//---------------------------------------------------------------------------------------------------------------
//
//  HAUD 2026.10.25
//
//  - ExternControl
//
//    - this is the main switchboard
//
//    - Transport abstractions are called here:
//    --------------------------------------------
//    - top level transport abstractions
//      - Instances contain the required transport logic
//      - Instances control their assigned ProcessCollector
//      - Instances are controlled in timer based application
//
//    - mid level transport abstractions
//      - StationCollectors and by extension ProcessCollectors
//      - Collectors are for gathering states and routing commands to ST_STATION_CTRL/STATE
//      - Collectors are configured during startup
//
//---------------------------------------------------------------------------------------------------------------
PROGRAM MAIN_APP
VAR
  eInitXtsTransport   AT %I*    : E_PROGRESS;   // initialization from XtsTransport PLC
  eInit               AT %Q*    : E_PROGRESS;   // local startup transmitted to TowerControl

  idx                           : UINT;
  nProcess                      : E_INSTANCE;

  // message pipeline(s) handling
  eMtrState,
  eMsgState                     : E_MESSAGE_STATE;
  eMtrProgress,
  eMsgProgress                  : E_PROGRESS;
  stMsg                         : ST_Message;
  //-------------------------------------------------------------------------------------------------------------
  tIdleWriteMotion              : TIME := T#5S;
  tIdleWriteApplication         : TIME := T#5S;
  tIdleWriteMetric              : TIME := T#5S;
  tonIdleWriteMotion            : Tc2_Standard.TON;
  tonIdleWriteApplication       : Tc2_Standard.TON;
  tonIdleWriteMetric            : Tc2_Standard.TON;
  //-------------------------------------------------------------------------------------------------------------
END_VAR

//#################################################################################################################
// Local time; used for timestamps
//#################################################################################################################
GVL_MSG_XTS.fbLocalTime();
GVL_MSG_XTS.sLocalTime                                            := GVL_MSG_XTS.fbLocalTime.LocalTimeString;
GVL_MSG_XTS.dtLocalTime                                           := GVL_MSG_XTS.fbLocalTime.LocalTime;
//-----------------------------------------------------------------------------------------------------------------
//-----------------------------------------------------------------------------------------------------------------
// check for Initialisation from XtsTransport first
//  - wait for XtsTransport to be fully started up
//-----------------------------------------------------------------------------------------------------------------
IF NOT (eInitXtsTransport = E_PROGRESS.PROGRESS_DONE) THEN eInit  := E_PROGRESS.PROGRESS_INVALID; RETURN; END_IF
//-----------------------------------------------------------------------------------------------------------------
//-----------------------------------------------------------------------------------------------------------------
// initialization for:
//  - configuring processes
//  - starting up of processes
//  - cross checking with the rest of your application
//-----------------------------------------------------------------------------------------------------------------
CASE eInit
OF
  E_PROGRESS.PROGRESS_INVALID:
    GVL_MSG_XTS.MetricsMessageCtrl.Cmd            := E_MESSAGE_CTRL.MSG_CTRL_INIT;
    eInit                                         := E_PROGRESS.PROGRESS_INIT;

  E_PROGRESS.PROGRESS_INIT:
    // init processes
    eInit                                         := E_PROGRESS.PROGRESS_BUSY;
    //-----------------------------------------------------------------------------
    //#############################################################################
    //-----------------------------------------------------------------------------
    GVL_APPLICATION.ProcessCollector[DISTRIBUTOR_INFEED].ProcessId            := DISTRIBUTOR_INFEED;
    GVL_APPLICATION.ProcessCollector[DISTRIBUTOR_INFEED].StationFirst         :=   142;
    GVL_APPLICATION.ProcessCollector[DISTRIBUTOR_INFEED].StationLast          :=   142;
    //-----------------------------------------------------------------------------
    GVL_APPLICATION.InstanceDistributorInfeed.ProcessId                       := DISTRIBUTOR_INFEED;
    GVL_APPLICATION.InstanceDistributorInfeed.ProcessTarget                   := PROCESS_INFEED;
    GVL_APPLICATION.InstanceDistributorInfeed.CheckPositionStart              :=  4500.0;
    GVL_APPLICATION.InstanceDistributorInfeed.CheckPositionEnd                :=  5600.0;
    //-----------------------------------------------------------------------------
    GVL_APPLICATION.InstanceDistributorInfeed.CollectorInterface              :=   GVL_APPLICATION.ItfProcessCollector;
    GVL_APPLICATION.InstanceDistributorInfeed.ProcessLinkedLists              :=   GVL_APPLICATION.ItfProcessList;
    GVL_APPLICATION.InstanceDistributorInfeed.InstanceCtrl                    REF= GVL_APPLICATION.InstanceCtrl;
    GVL_APPLICATION.InstanceDistributorInfeed.InstanceState                   REF= GVL_APPLICATION.InstanceState;
    GVL_APPLICATION.InstanceDistributorInfeed.MessageLevel                    :=   E_MessageType.eMessageError;

    //-----------------------------------------------------------------------------
    //#############################################################################
    //-----------------------------------------------------------------------------
    GVL_APPLICATION.ProcessCollector[PROCESS_INFEED].ProcessId                := PROCESS_INFEED;
    GVL_APPLICATION.ProcessCollector[PROCESS_INFEED].StationFirst             :=    20;
    GVL_APPLICATION.ProcessCollector[PROCESS_INFEED].StationLast              :=    35;
    //-----------------------------------------------------------------------------
    GVL_APPLICATION.InstanceInfeed.ProcessId                                  := PROCESS_INFEED;
    GVL_APPLICATION.InstanceInfeed.ProcessTarget                              := CONTINUOUS_CLEAN;
    GVL_APPLICATION.InstanceInfeed.CheckPositionStart                         :=  9750.0;
    GVL_APPLICATION.InstanceInfeed.CheckPositionEnd                           := 12100.0;
    //-----------------------------------------------------------------------------
    GVL_APPLICATION.InstanceInfeed.CollectorInterface                         :=   GVL_APPLICATION.ItfProcessCollector;
    GVL_APPLICATION.InstanceInfeed.ProcessLinkedLists                         :=   GVL_APPLICATION.ItfProcessList;
    GVL_APPLICATION.InstanceInfeed.InstanceCtrl                               REF= GVL_APPLICATION.InstanceCtrl;
    GVL_APPLICATION.InstanceInfeed.InstanceState                              REF= GVL_APPLICATION.InstanceState;
    GVL_APPLICATION.InstanceInfeed.MessageLevel                               :=   E_MessageType.eMessageError;

    //-----------------------------------------------------------------------------
    //#############################################################################
    //-----------------------------------------------------------------------------
    GVL_APPLICATION.ProcessCollector[CONTINUOUS_CLEAN].ProcessId              := CONTINUOUS_CLEAN;
    GVL_APPLICATION.ProcessCollector[CONTINUOUS_CLEAN].StationFirst           :=    37;
    GVL_APPLICATION.ProcessCollector[CONTINUOUS_CLEAN].StationLast            :=    37;
    //-----------------------------------------------------------------------------
    GVL_APPLICATION.InstanceCleaner.ProcessId                                 := CONTINUOUS_CLEAN;
    GVL_APPLICATION.InstanceCleaner.ProcessTarget                             := CONTINUOUS_SCAN;
    GVL_APPLICATION.InstanceCleaner.CheckPositionStart                        := 12850.0;
    GVL_APPLICATION.InstanceCleaner.CheckPositionEnd                          := 13000.0;
    //-----------------------------------------------------------------------------
    GVL_APPLICATION.InstanceCleaner.CollectorInterface                        :=   GVL_APPLICATION.ItfProcessCollector;
    GVL_APPLICATION.InstanceCleaner.ProcessLinkedLists                        :=   GVL_APPLICATION.ItfProcessList;
    GVL_APPLICATION.InstanceCleaner.InstanceCtrl                              REF= GVL_APPLICATION.InstanceCtrl;
    GVL_APPLICATION.InstanceCleaner.InstanceState                             REF= GVL_APPLICATION.InstanceState;

    //-----------------------------------------------------------------------------
    //#############################################################################
    //-----------------------------------------------------------------------------
    GVL_APPLICATION.ProcessCollector[CONTINUOUS_SCAN].ProcessId               := CONTINUOUS_SCAN;
    GVL_APPLICATION.ProcessCollector[CONTINUOUS_SCAN].StationFirst            :=    38;
    GVL_APPLICATION.ProcessCollector[CONTINUOUS_SCAN].StationLast             :=    38;
    //-----------------------------------------------------------------------------
    GVL_APPLICATION.InstanceScanner.ProcessId                                 := CONTINUOUS_SCAN;
    GVL_APPLICATION.InstanceScanner.ProcessTarget                             := CONTINUOUS_CAMERA;
    GVL_APPLICATION.InstanceScanner.CheckPositionStart                        := 13900.0;
    GVL_APPLICATION.InstanceScanner.CheckPositionEnd                          := 14100.0;
    //-----------------------------------------------------------------------------
    GVL_APPLICATION.InstanceScanner.CollectorInterface                        :=   GVL_APPLICATION.ItfProcessCollector;
    GVL_APPLICATION.InstanceScanner.ProcessLinkedLists                        :=   GVL_APPLICATION.ItfProcessList;
    GVL_APPLICATION.InstanceScanner.InstanceCtrl                              REF= GVL_APPLICATION.InstanceCtrl;
    GVL_APPLICATION.InstanceScanner.InstanceState                             REF= GVL_APPLICATION.InstanceState;

    //-----------------------------------------------------------------------------
    //#############################################################################
    //-----------------------------------------------------------------------------
    GVL_APPLICATION.ProcessCollector[CONTINUOUS_CAMERA].ProcessId             := CONTINUOUS_CAMERA;
    GVL_APPLICATION.ProcessCollector[CONTINUOUS_CAMERA].StationFirst          :=    39;
    GVL_APPLICATION.ProcessCollector[CONTINUOUS_CAMERA].StationLast           :=    39;
    //-----------------------------------------------------------------------------
    GVL_APPLICATION.InstanceCamera.ProcessId                                  := CONTINUOUS_CAMERA;
    GVL_APPLICATION.InstanceCamera.ProcessTarget                              := DISTRIBUTOR_ASSEMBLY_01;
    GVL_APPLICATION.InstanceCamera.CheckPositionStart                         := 14200.0;
    GVL_APPLICATION.InstanceCamera.CheckPositionEnd                           := 14400.0;
    //-----------------------------------------------------------------------------
    GVL_APPLICATION.InstanceCamera.CollectorInterface                         :=   GVL_APPLICATION.ItfProcessCollector;
    GVL_APPLICATION.InstanceCamera.ProcessLinkedLists                         :=   GVL_APPLICATION.ItfProcessList;
    GVL_APPLICATION.InstanceCamera.InstanceCtrl                               REF= GVL_APPLICATION.InstanceCtrl;
    GVL_APPLICATION.InstanceCamera.InstanceState                              REF= GVL_APPLICATION.InstanceState;

    //-----------------------------------------------------------------------------
    //#############################################################################
    //-----------------------------------------------------------------------------
    GVL_APPLICATION.ProcessCollector[DISTRIBUTOR_ASSEMBLY_01].ProcessId       := DISTRIBUTOR_ASSEMBLY_01;
    GVL_APPLICATION.ProcessCollector[DISTRIBUTOR_ASSEMBLY_01].StationFirst    :=    40;
    GVL_APPLICATION.ProcessCollector[DISTRIBUTOR_ASSEMBLY_01].StationLast     :=    40;
    //-----------------------------------------------------------------------------
    GVL_APPLICATION.InstanceDistributorAssembly_01.ProcessId                  := DISTRIBUTOR_ASSEMBLY_01;
    GVL_APPLICATION.InstanceDistributorAssembly_01.ProcessTarget              := PROCESS_ASSEMBLY_01;
    GVL_APPLICATION.InstanceDistributorAssembly_01.CheckPositionStart         := 14400.0;
    GVL_APPLICATION.InstanceDistributorAssembly_01.CheckPositionEnd           := 17500.0;
    //-----------------------------------------------------------------------------
    GVL_APPLICATION.InstanceDistributorAssembly_01.CollectorInterface         :=   GVL_APPLICATION.ItfProcessCollector;
    GVL_APPLICATION.InstanceDistributorAssembly_01.ProcessLinkedLists         :=   GVL_APPLICATION.ItfProcessList;
    GVL_APPLICATION.InstanceDistributorAssembly_01.InstanceCtrl               REF= GVL_APPLICATION.InstanceCtrl;
    GVL_APPLICATION.InstanceDistributorAssembly_01.InstanceState              REF= GVL_APPLICATION.InstanceState;

    //-----------------------------------------------------------------------------
    //#############################################################################
    //-----------------------------------------------------------------------------
    GVL_APPLICATION.ProcessCollector[PROCESS_ASSEMBLY_01].ProcessId           := PROCESS_ASSEMBLY_01;
    GVL_APPLICATION.ProcessCollector[PROCESS_ASSEMBLY_01].StationFirst        :=    41;
    GVL_APPLICATION.ProcessCollector[PROCESS_ASSEMBLY_01].StationLast         :=    56;
    //-----------------------------------------------------------------------------
    GVL_APPLICATION.InstanceAssembly_01.ProcessId                             := PROCESS_ASSEMBLY_01;
    GVL_APPLICATION.InstanceAssembly_01.ProcessTarget                         := DISTRIBUTOR_ASSEMBLY_02;
    GVL_APPLICATION.InstanceAssembly_01.CheckPositionStart                    := 14400.0;
    GVL_APPLICATION.InstanceAssembly_01.CheckPositionEnd                      := 17500.0;
    //-----------------------------------------------------------------------------
    GVL_APPLICATION.InstanceAssembly_01.CollectorInterface                    :=   GVL_APPLICATION.ItfProcessCollector;
    GVL_APPLICATION.InstanceAssembly_01.ProcessLinkedLists                    :=   GVL_APPLICATION.ItfProcessList;
    GVL_APPLICATION.InstanceAssembly_01.InstanceCtrl                          REF= GVL_APPLICATION.InstanceCtrl;
    GVL_APPLICATION.InstanceAssembly_01.InstanceState                         REF= GVL_APPLICATION.InstanceState;

    //-----------------------------------------------------------------------------
    //#############################################################################
    //-----------------------------------------------------------------------------
    GVL_APPLICATION.ProcessCollector[DISTRIBUTOR_ASSEMBLY_02].ProcessId       := DISTRIBUTOR_ASSEMBLY_02;
    GVL_APPLICATION.ProcessCollector[DISTRIBUTOR_ASSEMBLY_02].StationFirst    :=    57;
    GVL_APPLICATION.ProcessCollector[DISTRIBUTOR_ASSEMBLY_02].StationLast     :=    57;
    //-----------------------------------------------------------------------------
    GVL_APPLICATION.InstanceDistributorAssembly_02.ProcessId                  := DISTRIBUTOR_ASSEMBLY_02;
    GVL_APPLICATION.InstanceDistributorAssembly_02.ProcessTarget              := PROCESS_ASSEMBLY_02;
    GVL_APPLICATION.InstanceDistributorAssembly_02.CheckPositionStart         := 17500.0;
    GVL_APPLICATION.InstanceDistributorAssembly_02.CheckPositionEnd           := 18100.0;
    //-----------------------------------------------------------------------------
    GVL_APPLICATION.InstanceDistributorAssembly_02.CollectorInterface         :=   GVL_APPLICATION.ItfProcessCollector;
    GVL_APPLICATION.InstanceDistributorAssembly_02.ProcessLinkedLists         :=   GVL_APPLICATION.ItfProcessList;
    GVL_APPLICATION.InstanceDistributorAssembly_02.InstanceCtrl               REF= GVL_APPLICATION.InstanceCtrl;
    GVL_APPLICATION.InstanceDistributorAssembly_02.InstanceState              REF= GVL_APPLICATION.InstanceState;

    //-----------------------------------------------------------------------------
    //#############################################################################
    //-----------------------------------------------------------------------------
    GVL_APPLICATION.ProcessCollector[PROCESS_ASSEMBLY_02].ProcessId           := PROCESS_ASSEMBLY_02;
    GVL_APPLICATION.ProcessCollector[PROCESS_ASSEMBLY_02].StationFirst        :=    58;
    GVL_APPLICATION.ProcessCollector[PROCESS_ASSEMBLY_02].StationLast         :=    67;
    //-----------------------------------------------------------------------------
    GVL_APPLICATION.InstanceAssembly_02.ProcessId                             := PROCESS_ASSEMBLY_02;
    GVL_APPLICATION.InstanceAssembly_02.ProcessTarget                         := DISTRIBUTOR_ASSEMBLY_TEST;
    GVL_APPLICATION.InstanceAssembly_02.CheckPositionStart                    := 19400.0;
    GVL_APPLICATION.InstanceAssembly_02.CheckPositionEnd                      := 20750.0;
    //-----------------------------------------------------------------------------
    GVL_APPLICATION.InstanceAssembly_02.CollectorInterface                    :=   GVL_APPLICATION.ItfProcessCollector;
    GVL_APPLICATION.InstanceAssembly_02.ProcessLinkedLists                    :=   GVL_APPLICATION.ItfProcessList;
    GVL_APPLICATION.InstanceAssembly_02.InstanceCtrl                          REF= GVL_APPLICATION.InstanceCtrl;
    GVL_APPLICATION.InstanceAssembly_02.InstanceState                         REF= GVL_APPLICATION.InstanceState;

    //-----------------------------------------------------------------------------
    //#############################################################################
    //-----------------------------------------------------------------------------
    GVL_APPLICATION.ProcessCollector[DISTRIBUTOR_ASSEMBLY_TEST].ProcessId     := DISTRIBUTOR_ASSEMBLY_TEST;
    GVL_APPLICATION.ProcessCollector[DISTRIBUTOR_ASSEMBLY_TEST].StationFirst  :=    70;
    GVL_APPLICATION.ProcessCollector[DISTRIBUTOR_ASSEMBLY_TEST].StationLast   :=    70;
    //-----------------------------------------------------------------------------
    GVL_APPLICATION.InstanceDistributorAssemblyTest.ProcessId                 := DISTRIBUTOR_ASSEMBLY_TEST;
    GVL_APPLICATION.InstanceDistributorAssemblyTest.ProcessTarget             := PROCESS_ASSEMBLY_TEST;
    GVL_APPLICATION.InstanceDistributorAssemblyTest.CheckPositionStart        := 20600.0;
    GVL_APPLICATION.InstanceDistributorAssemblyTest.CheckPositionEnd          := 21400.0;
    //-----------------------------------------------------------------------------
    GVL_APPLICATION.InstanceDistributorAssemblyTest.CollectorInterface        :=   GVL_APPLICATION.ItfProcessCollector;
    GVL_APPLICATION.InstanceDistributorAssemblyTest.ProcessLinkedLists        :=   GVL_APPLICATION.ItfProcessList;
    GVL_APPLICATION.InstanceDistributorAssemblyTest.InstanceCtrl              REF= GVL_APPLICATION.InstanceCtrl;
    GVL_APPLICATION.InstanceDistributorAssemblyTest.InstanceState             REF= GVL_APPLICATION.InstanceState;

    //-----------------------------------------------------------------------------
    //#############################################################################
    //-----------------------------------------------------------------------------
    GVL_APPLICATION.ProcessCollector[PROCESS_ASSEMBLY_TEST].ProcessId         := PROCESS_ASSEMBLY_TEST;
    GVL_APPLICATION.ProcessCollector[PROCESS_ASSEMBLY_TEST].StationFirst      :=    71;
    GVL_APPLICATION.ProcessCollector[PROCESS_ASSEMBLY_TEST].StationLast       :=    86;
    //-----------------------------------------------------------------------------
    GVL_APPLICATION.InstanceAssemblyTest.ProcessId                            := PROCESS_ASSEMBLY_TEST;
    GVL_APPLICATION.InstanceAssemblyTest.ProcessTarget                        := DISTRIBUTOR_CAMERA;
    GVL_APPLICATION.InstanceAssemblyTest.CheckPositionStart                   := 21400.0;
    GVL_APPLICATION.InstanceAssemblyTest.CheckPositionEnd                     := 23000.0;
    //-----------------------------------------------------------------------------
    GVL_APPLICATION.InstanceAssemblyTest.CollectorInterface                   :=   GVL_APPLICATION.ItfProcessCollector;
    GVL_APPLICATION.InstanceAssemblyTest.ProcessLinkedLists                   :=   GVL_APPLICATION.ItfProcessList;
    GVL_APPLICATION.InstanceAssemblyTest.InstanceCtrl                         REF= GVL_APPLICATION.InstanceCtrl;
    GVL_APPLICATION.InstanceAssemblyTest.InstanceState                        REF= GVL_APPLICATION.InstanceState;

    //-----------------------------------------------------------------------------
    //#############################################################################
    //-----------------------------------------------------------------------------
    GVL_APPLICATION.ProcessCollector[DISTRIBUTOR_CAMERA].ProcessId            := DISTRIBUTOR_CAMERA;
    GVL_APPLICATION.ProcessCollector[DISTRIBUTOR_CAMERA].StationFirst         :=    91;
    GVL_APPLICATION.ProcessCollector[DISTRIBUTOR_CAMERA].StationLast          :=    91;
    //-----------------------------------------------------------------------------
    GVL_APPLICATION.InstanceAssemblyCameraInfeed.ProcessId                    := DISTRIBUTOR_CAMERA;
    GVL_APPLICATION.InstanceAssemblyCameraInfeed.ProcessTarget                := CONTINUOUS_ASSEMBLY_CAMERA;
    GVL_APPLICATION.InstanceAssemblyCameraInfeed.CheckPositionStart           := 22800.0;
    GVL_APPLICATION.InstanceAssemblyCameraInfeed.CheckPositionEnd             := 23500.0;
    //-----------------------------------------------------------------------------
    GVL_APPLICATION.InstanceAssemblyCameraInfeed.CollectorInterface           :=   GVL_APPLICATION.ItfProcessCollector;
    GVL_APPLICATION.InstanceAssemblyCameraInfeed.ProcessLinkedLists           :=   GVL_APPLICATION.ItfProcessList;
    GVL_APPLICATION.InstanceAssemblyCameraInfeed.InstanceCtrl                 REF= GVL_APPLICATION.InstanceCtrl;
    GVL_APPLICATION.InstanceAssemblyCameraInfeed.InstanceState                REF= GVL_APPLICATION.InstanceState;

    //-----------------------------------------------------------------------------
    //#############################################################################
    //-----------------------------------------------------------------------------
    GVL_APPLICATION.ProcessCollector[CONTINUOUS_ASSEMBLY_CAMERA].ProcessId    := CONTINUOUS_ASSEMBLY_CAMERA;
    GVL_APPLICATION.ProcessCollector[CONTINUOUS_ASSEMBLY_CAMERA].StationFirst :=    95;
    GVL_APPLICATION.ProcessCollector[CONTINUOUS_ASSEMBLY_CAMERA].StationLast  :=    95;
    //-----------------------------------------------------------------------------
    GVL_APPLICATION.InstanceAssemblyCameraOutfeed.ProcessId                   := CONTINUOUS_ASSEMBLY_CAMERA;
    GVL_APPLICATION.InstanceAssemblyCameraOutfeed.ProcessTarget               := DISTRIBUTOR_OUTFEED;
    GVL_APPLICATION.InstanceAssemblyCameraOutfeed.CheckPositionStart          := 24000.0;
    GVL_APPLICATION.InstanceAssemblyCameraOutfeed.CheckPositionEnd            := 24100.0;
    //-----------------------------------------------------------------------------
    GVL_APPLICATION.InstanceAssemblyCameraOutfeed.CollectorInterface          :=   GVL_APPLICATION.ItfProcessCollector;
    GVL_APPLICATION.InstanceAssemblyCameraOutfeed.ProcessLinkedLists          :=   GVL_APPLICATION.ItfProcessList;
    GVL_APPLICATION.InstanceAssemblyCameraOutfeed.InstanceCtrl                REF= GVL_APPLICATION.InstanceCtrl;
    GVL_APPLICATION.InstanceAssemblyCameraOutfeed.InstanceState               REF= GVL_APPLICATION.InstanceState;

    //-----------------------------------------------------------------------------
    //#############################################################################
    //-----------------------------------------------------------------------------
    GVL_APPLICATION.ProcessCollector[DISTRIBUTOR_OUTFEED].ProcessId           := DISTRIBUTOR_OUTFEED;
    GVL_APPLICATION.ProcessCollector[DISTRIBUTOR_OUTFEED].StationFirst        :=   119;
    GVL_APPLICATION.ProcessCollector[DISTRIBUTOR_OUTFEED].StationLast         :=   119;
    //-----------------------------------------------------------------------------
    GVL_APPLICATION.InstanceDistributorOutfeed.ProcessId                      := DISTRIBUTOR_OUTFEED;
    GVL_APPLICATION.InstanceDistributorOutfeed.ProcessTarget                  := PROCESS_OUTFEED;
    GVL_APPLICATION.InstanceDistributorOutfeed.CheckPositionStart             := 24000.0;
    GVL_APPLICATION.InstanceDistributorOutfeed.CheckPositionEnd               := 27500.0;
    //-----------------------------------------------------------------------------
    GVL_APPLICATION.InstanceDistributorOutfeed.CollectorInterface             :=   GVL_APPLICATION.ItfProcessCollector;
    GVL_APPLICATION.InstanceDistributorOutfeed.ProcessLinkedLists             :=   GVL_APPLICATION.ItfProcessList;
    GVL_APPLICATION.InstanceDistributorOutfeed.InstanceCtrl                   REF= GVL_APPLICATION.InstanceCtrl;
    GVL_APPLICATION.InstanceDistributorOutfeed.InstanceState                  REF= GVL_APPLICATION.InstanceState;

    //-----------------------------------------------------------------------------
    //#############################################################################
    //-----------------------------------------------------------------------------
    GVL_APPLICATION.ProcessCollector[PROCESS_OUTFEED].ProcessId               := PROCESS_OUTFEED;
    GVL_APPLICATION.ProcessCollector[PROCESS_OUTFEED].StationFirst            :=   120;
    GVL_APPLICATION.ProcessCollector[PROCESS_OUTFEED].StationLast             :=   133;
    //-----------------------------------------------------------------------------
    GVL_APPLICATION.InstanceOutfeed.ProcessId                                 := PROCESS_OUTFEED;
    GVL_APPLICATION.InstanceOutfeed.ProcessTarget                             := DISTRIBUTOR_WPC_CLEAN;
    GVL_APPLICATION.InstanceOutfeed.CheckPositionStart                        := 24500.0;
    GVL_APPLICATION.InstanceOutfeed.CheckPositionEnd                          := 27500.0;
    //-----------------------------------------------------------------------------
    GVL_APPLICATION.InstanceOutfeed.CollectorInterface                        :=   GVL_APPLICATION.ItfProcessCollector;
    GVL_APPLICATION.InstanceOutfeed.ProcessLinkedLists                        :=   GVL_APPLICATION.ItfProcessList;
    GVL_APPLICATION.InstanceOutfeed.InstanceCtrl                              REF= GVL_APPLICATION.InstanceCtrl;
    GVL_APPLICATION.InstanceOutfeed.InstanceState                             REF= GVL_APPLICATION.InstanceState;

    //-----------------------------------------------------------------------------
    //#############################################################################
    //-----------------------------------------------------------------------------
    GVL_APPLICATION.ProcessCollector[DISTRIBUTOR_WPC_CLEAN].ProcessId         := DISTRIBUTOR_WPC_CLEAN;
    GVL_APPLICATION.ProcessCollector[DISTRIBUTOR_WPC_CLEAN].StationFirst      :=   140;
    GVL_APPLICATION.ProcessCollector[DISTRIBUTOR_WPC_CLEAN].StationLast       :=   140;
    //-----------------------------------------------------------------------------
    GVL_APPLICATION.InstanceDistributorWpcClean.ProcessId                     := DISTRIBUTOR_WPC_CLEAN;
    GVL_APPLICATION.InstanceDistributorWpcClean.ProcessTarget                 := CONTINUOUS_WPC_CLEAN;
    GVL_APPLICATION.InstanceDistributorWpcClean.CheckPositionStart            := 27970.0;
    GVL_APPLICATION.InstanceDistributorWpcClean.CheckPositionEnd              :=  1250.0;
    //-----------------------------------------------------------------------------
    GVL_APPLICATION.InstanceDistributorWpcClean.CollectorInterface            :=   GVL_APPLICATION.ItfProcessCollector;
    GVL_APPLICATION.InstanceDistributorWpcClean.ProcessLinkedLists            :=   GVL_APPLICATION.ItfProcessList;
    GVL_APPLICATION.InstanceDistributorWpcClean.InstanceCtrl                  REF= GVL_APPLICATION.InstanceCtrl;
    GVL_APPLICATION.InstanceDistributorWpcClean.InstanceState                 REF= GVL_APPLICATION.InstanceState;

    //-----------------------------------------------------------------------------
    //#############################################################################
    //-----------------------------------------------------------------------------
    GVL_APPLICATION.ProcessCollector[CONTINUOUS_WPC_CLEAN].ProcessId          := CONTINUOUS_WPC_CLEAN;
    GVL_APPLICATION.ProcessCollector[CONTINUOUS_WPC_CLEAN].StationFirst       :=   141;
    GVL_APPLICATION.ProcessCollector[CONTINUOUS_WPC_CLEAN].StationLast        :=   141;
    //-----------------------------------------------------------------------------
    GVL_APPLICATION.InstanceWpcClean.ProcessId                                := CONTINUOUS_WPC_CLEAN;
    GVL_APPLICATION.InstanceWpcClean.ProcessTarget                            := DISTRIBUTOR_INFEED;
    GVL_APPLICATION.InstanceWpcClean.CheckPositionStart                       :=  3950.0;
    GVL_APPLICATION.InstanceWpcClean.CheckPositionEnd                         :=  4100.0;
    //-----------------------------------------------------------------------------
    GVL_APPLICATION.InstanceWpcClean.CollectorInterface                       :=   GVL_APPLICATION.ItfProcessCollector;
    GVL_APPLICATION.InstanceWpcClean.ProcessLinkedLists                       :=   GVL_APPLICATION.ItfProcessList;
    GVL_APPLICATION.InstanceWpcClean.InstanceCtrl                             REF= GVL_APPLICATION.InstanceCtrl;
    GVL_APPLICATION.InstanceWpcClean.InstanceState                            REF= GVL_APPLICATION.InstanceState;


  E_PROGRESS.PROGRESS_BUSY:
    // init the conductor
    GVL_APPLICATION.ConductorCtrl.Cmd             := E_INSTANCE_CMD.INIT;
    // init the instances
    idx                                           := 1;
    memset(ADR(GVL_APPLICATION.InstanceCtrl), 0, SIZEOF(GVL_APPLICATION.InstanceCtrl));
    eInit                                         := E_PROGRESS.PROGRESS_PREPARE;

  E_PROGRESS.PROGRESS_PREPARE:
    GVL_APPLICATION.InstanceCtrl[idx].Cmd         := E_INSTANCE_CMD.INIT;

    IF (GVL_APPLICATION.InstanceState[idx].ProcessState   = E_INSTANCE_STATE.DISABLED)
    THEN
      IF (GVL_APPLICATION.InstanceState[idx].ProcessProgress = E_PROGRESS.PROGRESS_BUSY)
      THEN
        GVL_APPLICATION.InstanceCtrl[idx].Cmd     := E_INSTANCE_CMD.DISABLE;
        eInit                                     := E_PROGRESS.PROGRESS_STARTUP;
      END_IF
    END_IF


  E_PROGRESS.PROGRESS_STARTUP:
    IF NOT (idx < GVL_APPLICATION.MAX_PROCESS)
    THEN
      eInit                                       := E_PROGRESS.PROGRESS_CHECK;
    ELSE
      idx                                         := idx + 1;
      eInit                                       := E_PROGRESS.PROGRESS_PREPARE;
    END_IF

  E_PROGRESS.PROGRESS_CHECK:
    GVL_APPLICATION.ConductorCtrl.Cmd             := E_INSTANCE_CMD.ENABLE;
    eInit                                         := E_PROGRESS.PROGRESS_OCCUPIED;

  E_PROGRESS.PROGRESS_OCCUPIED:
    eInit                                         := E_PROGRESS.PROGRESS_WORKING;

  E_PROGRESS.PROGRESS_WORKING:
    eInit                                         := E_PROGRESS.PROGRESS_DONE;
END_CASE
//-----------------------------------------------------------------------------------------------------------------
//-----------------------------------------------------------------------------------------------------------------
//-----------------------------------------------------------------------------------------------------------------
//-----------------------------------------------------------------------------------------------------------------
// /assign dataflow
//-----------------------------------------------------------------------------------------------------------------
//-----------------------------------------------------------------------------------------------------------------
//  - The YardMaster
//-----------------------------------------------------------------------------------------------------------------
GVL_APPLICATION.YardMaster.Ctrl                               REF= GVL_APPLICATION.YardControl;
GVL_APPLICATION.YardMaster.State                              REF= GVL_APPLICATION.YardState;

GVL_APPLICATION.YardMaster.XtsTransportCtrl                   REF= GVL_XTS.XtsTransportCtrl;
GVL_APPLICATION.YardMaster.XtsTransportState                  REF= GVL_XTS.XtsTransportState;

GVL_APPLICATION.YardMaster.CollectorInterfaces                :=   GVL_APPLICATION.ItfProcessCollector;
GVL_APPLICATION.YardMaster.TicketList                         :=   GVL_APPLICATION.TicketList;
GVL_APPLICATION.YardMaster();
//-----------------------------------------------------------------------------------------------------------------
//  - ProcessCollectors
//-----------------------------------------------------------------------------------------------------------------
FOR nProcess := 1 TO MAX_PROCESS
DO
  GVL_APPLICATION.ItfProcessList[nProcess]                    :=   GVL_APPLICATION.ProcessList[nProcess];
  GVL_APPLICATION.ItfProcessCollector[nProcess]               :=   GVL_APPLICATION.ProcessCollector[nProcess];

  GVL_APPLICATION.ProcessCollector[nProcess].MessageLevel     :=   GVL_MSG_XTS.MessageLevelProcess[nProcess];
  GVL_APPLICATION.ProcessCollector[nProcess].MoverInfo        REF= GVL_XTS.MoverInfo;
  GVL_APPLICATION.ProcessCollector[nProcess].StationCtrl      REF= GVL_XTS.StationCtrl;
  GVL_APPLICATION.ProcessCollector[nProcess].StationState     REF= GVL_XTS.StationState;
  GVL_APPLICATION.ProcessCollector[nProcess].Cycle();
END_FOR
//-----------------------------------------------------------------------------------------------------------------
//-----------------------------------------------------------------------------------------------------------------
// cyclic TicketList as inbox
//-----------------------------------------------------------------------------------------------------------------
//-----------------------------------------------------------------------------------------------------------------
GVL_APPLICATION.TicketControl.ItfList                         :=   GVL_APPLICATION.TicketList;
GVL_APPLICATION.TicketControl.Ctrl                            REF= GVL_APPLICATION.TicketListControl;
GVL_APPLICATION.TicketControl.State                           REF= GVL_APPLICATION.TicketListState;
GVL_APPLICATION.TicketControl.NodeDataInput                   REF= GVL_APPLICATION.TicketListDataInput;
GVL_APPLICATION.TicketControl.NodeDataOutput                  REF= GVL_APPLICATION.TicketListDataOutput;
GVL_APPLICATION.TicketControl();
//-----------------------------------------------------------------------------------------------------------------
//-----------------------------------------------------------------------------------------------------------------
// Conductor
//-----------------------------------------------------------------------------------------------------------------
//-----------------------------------------------------------------------------------------------------------------
GVL_APPLICATION.ProcessConductor.ProcessLinkedLists           :=   GVL_APPLICATION.ItfProcessList;
GVL_APPLICATION.ProcessConductor.TicketLinkedList             :=   GVL_APPLICATION.TicketList;
GVL_APPLICATION.ProcessConductor.Ctrl                         REF= GVL_APPLICATION.ConductorCtrl;
GVL_APPLICATION.ProcessConductor.State                        REF= GVL_APPLICATION.ConductorState;
GVL_APPLICATION.ProcessConductor();
//-----------------------------------------------------------------------------------------------------------------
//-----------------------------------------------------------------------------------------------------------------
// Instance calls
//-----------------------------------------------------------------------------------------------------------------
//-----------------------------------------------------------------------------------------------------------------
GVL_APPLICATION.InstanceWpcClean();
GVL_APPLICATION.InstanceDistributorWpcClean();
GVL_APPLICATION.InstanceOutfeed();
GVL_APPLICATION.InstanceDistributorOutfeed();
GVL_APPLICATION.InstanceAssemblyCameraOutfeed();
GVL_APPLICATION.InstanceAssemblyCameraInfeed();
GVL_APPLICATION.InstanceAssemblyTest();
GVL_APPLICATION.InstanceDistributorAssemblyTest();
GVL_APPLICATION.InstanceAssembly_02();
GVL_APPLICATION.InstanceDistributorAssembly_02();
GVL_APPLICATION.InstanceAssembly_01();
GVL_APPLICATION.InstanceDistributorAssembly_01();
GVL_APPLICATION.InstanceCamera();
GVL_APPLICATION.InstanceScanner();
GVL_APPLICATION.InstanceCleaner();
GVL_APPLICATION.InstanceInfeed();
GVL_APPLICATION.InstanceDistributorInfeed();
//-----------------------------------------------------------------------------------------------------------------
//-----------------------------------------------------------------------------------------------------------------
//#################################################################################################################
//  /logging
//    - all life is problem solving
//#################################################################################################################
GVL_MSG_XTS.TransportMessageData.Ctrl               REF= GVL_MSG_XTS.TransportMessageCtrl;
GVL_MSG_XTS.TransportMessageData.State              REF= GVL_MSG_XTS.TransportMessageState;
GVL_MSG_XTS.TransportMessageData.MessageIndex       REF= GVL_MSG_XTS.MessageTransportIndex;
GVL_MSG_XTS.TransportMessageData.ErrorIndex         REF= GVL_MSG_XTS.MessageTransportError;
GVL_MSG_XTS.TransportMessageData.DirRoot            :=   ADR(GVL_MSG_XTS.LOG_DIR);
GVL_MSG_XTS.TransportMessageData.FileRoot           :=   ADR(GVL_MSG_XTS.LOG_FILE);
GVL_MSG_XTS.TransportMessageData.MsgList            :=   ADR(GVL_MSG_XTS.TransportMessages);
GVL_MSG_XTS.TransportMessageData.LocalTime          :=   ADR(GVL_MSG_XTS.dtLocalTime);
GVL_MSG_XTS.TransportMessageData();
eMsgState                                       :=   f_GetState   (GVL_MSG_XTS.TransportMessageState.State);
eMsgProgress                                    :=   f_GetProgress(GVL_MSG_XTS.TransportMessageState.State);

CASE eMsgState
OF
  E_MESSAGE_STATE.MSG_STATE_NULL:
    CASE eMsgProgress
    OF
      E_PROGRESS.PROGRESS_INVALID,
      E_PROGRESS.PROGRESS_DONE:
        IF (GVL_MSG_XTS.MessageTransportIndex > GVL_MSG_XTS.MAX_MESSAGE/101) OR
           (GVL_MSG_XTS.MessageTransportError > 0)
        THEN
          GVL_MSG_XTS.TransportMessageCtrl.Cmd      := E_MESSAGE_CTRL.MSG_CTRL_WRITE;
        ELSE
          tonIdleWriteMotion(IN := TRUE, PT:= tIdleWriteMotion);
          IF (tonIdleWriteMotion.Q)
          THEN
            GVL_MSG_XTS.TransportMessageCtrl.Cmd    := E_MESSAGE_CTRL.MSG_CTRL_WRITE;
          END_IF
        END_IF
    END_CASE

  E_MESSAGE_STATE.MSG_STATE_WRITE:
    CASE eMsgProgress
    OF
      E_PROGRESS.PROGRESS_ERROR,
      E_PROGRESS.PROGRESS_DONE:
          tonIdleWriteMotion(IN := FALSE, PT:= tIdleWriteMotion);
        GVL_MSG_XTS.TransportMessageCtrl.Cmd        := E_MESSAGE_CTRL.MSG_CTRL_NULL;
    END_CASE

ELSE
    CASE eMsgProgress
    OF
      E_PROGRESS.PROGRESS_DONE:
          tonIdleWriteMotion(IN := FALSE, PT:= tIdleWriteMotion);
        GVL_MSG_XTS.TransportMessageCtrl.Cmd        := E_MESSAGE_CTRL.MSG_CTRL_NULL;
    END_CASE
END_CASE
//#################################################################################################################
// /application logging
//#################################################################################################################
GVL_MSG_XTS.ApplicationMessageData.Ctrl                         REF= GVL_MSG_XTS.ApplicationMessageCtrl;
GVL_MSG_XTS.ApplicationMessageData.State                        REF= GVL_MSG_XTS.ApplicationMessageState;

GVL_MSG_XTS.ApplicationMessageData.MessageIndex                 REF= GVL_MSG_XTS.MessageApplicationIndex;
GVL_MSG_XTS.ApplicationMessageData.ErrorIndex                   REF= GVL_MSG_XTS.MessageApplicationError;

GVL_MSG_XTS.ApplicationMessageData.DirRoot                      :=   ADR(GVL_MSG_XTS.LOG_DIR);
GVL_MSG_XTS.ApplicationMessageData.FileRoot                     :=   ADR(GVL_MSG_XTS.LOG_FILE_APP);
GVL_MSG_XTS.ApplicationMessageData.MsgList                      :=   ADR(GVL_MSG_XTS.ApplicationMessages);
GVL_MSG_XTS.ApplicationMessageData.LocalTime                    :=   ADR(GVL_MSG_XTS.dtLocalTime);

GVL_MSG_XTS.ApplicationMessageData();

eMsgState                                       := f_GetState   (GVL_MSG_XTS.ApplicationMessageState.State);
eMsgProgress                                    := f_GetProgress(GVL_MSG_XTS.ApplicationMessageState.State);


CASE eMsgState
OF
  E_MESSAGE_STATE.MSG_STATE_NULL:
    CASE eMsgProgress
    OF
      E_PROGRESS.PROGRESS_INVALID:
        IF (GVL_MSG_XTS.MessageApplicationIndex > GVL_MSG_XTS.MAX_MESSAGE/13) OR
           (GVL_MSG_XTS.MessageApplicationError > 0)
        THEN
          GVL_MSG_XTS.ApplicationMessageCtrl.Cmd                := E_MESSAGE_CTRL.MSG_CTRL_WRITE;
        ELSE
          tonIdleWriteApplication(IN := TRUE, PT:= tIdleWriteApplication);
          IF (tonIdleWriteApplication.Q)
          THEN
            GVL_MSG_XTS.ApplicationMessageCtrl.Cmd              := E_MESSAGE_CTRL.MSG_CTRL_WRITE;
          END_IF
        END_IF
    END_CASE

  E_MESSAGE_STATE.MSG_STATE_WRITE:
    CASE eMsgProgress
    OF
      E_PROGRESS.PROGRESS_ERROR,
      E_PROGRESS.PROGRESS_DONE:
        tonIdleWriteApplication(IN := FALSE, PT:= tIdleWriteApplication);
        GVL_MSG_XTS.ApplicationMessageCtrl.Cmd                  := E_MESSAGE_CTRL.MSG_CTRL_NULL;
    END_CASE

ELSE
    CASE eMsgProgress
    OF
      E_PROGRESS.PROGRESS_DONE:
        tonIdleWriteApplication(IN := FALSE, PT:= tIdleWriteApplication);
        GVL_MSG_XTS.ApplicationMessageCtrl.Cmd                  := E_MESSAGE_CTRL.MSG_CTRL_NULL;
    END_CASE
END_CASE
//#################################################################################################################
// logging/
//#################################################################################################################
//#################################################################################################################
//  /Transport Metrics
//#################################################################################################################
GVL_MSG_XTS.MetricsMessageData.Ctrl                             REF= GVL_MSG_XTS.MetricsMessageCtrl;
GVL_MSG_XTS.MetricsMessageData.State                            REF= GVL_MSG_XTS.MetricsMessageState;

GVL_MSG_XTS.MetricsMessageData.MessageIndex                     REF= GVL_MSG_XTS.MessageMetricsIndex;
GVL_MSG_XTS.MetricsMessageData.ErrorIndex                       REF= GVL_MSG_XTS.MessageMetricsError;

GVL_MSG_XTS.MetricsMessageData.DirRoot                          :=   ADR(GVL_MSG_XTS.LOG_DIR);
GVL_MSG_XTS.MetricsMessageData.FileRoot                         :=   ADR(GVL_MSG_XTS.LOG_FILE_METRIC);
GVL_MSG_XTS.MetricsMessageData.MsgList                          :=   ADR(GVL_MSG_XTS.MetricsMessages);
GVL_MSG_XTS.MetricsMessageData.LocalTime                        :=   ADR(GVL_MSG_XTS.dtLocalTime);

GVL_MSG_XTS.MetricsMessageData();

eMtrState                                   := f_GetState   (GVL_MSG_XTS.MetricsMessageState.State);
eMtrProgress                                := f_GetProgress(GVL_MSG_XTS.MetricsMessageState.State);

CASE eMtrState
OF
  E_MESSAGE_STATE.MSG_STATE_NULL:
    CASE eMtrProgress
    OF
      E_PROGRESS.PROGRESS_INVALID:
        IF (GVL_MSG_XTS.MessageMetricsIndex > GVL_MSG_XTS.MAX_MESSAGE/5) OR
           (GVL_MSG_XTS.MessageMetricsError > 0)
        THEN
          GVL_MSG_XTS.MetricsMessageCtrl.Cmd                    := E_MESSAGE_CTRL.MSG_CTRL_WRITE;
        ELSE
          tonIdleWriteMetric(IN := TRUE, PT:= tIdleWriteMetric);
          IF (tonIdleWriteMetric.Q)
          THEN
            GVL_MSG_XTS.MetricsMessageCtrl.Cmd                  := E_MESSAGE_CTRL.MSG_CTRL_WRITE;
          END_IF
        END_IF
    END_CASE

  E_MESSAGE_STATE.MSG_STATE_WRITE:
    CASE eMtrProgress
    OF
      E_PROGRESS.PROGRESS_ERROR,
      E_PROGRESS.PROGRESS_DONE:
        tonIdleWriteMetric(IN := FALSE, PT:= tIdleWriteMetric);
        GVL_MSG_XTS.MetricsMessageCtrl.Cmd                      := E_MESSAGE_CTRL.MSG_CTRL_NULL;
    END_CASE
ELSE
    CASE eMtrProgress
    OF
      E_PROGRESS.PROGRESS_DONE:
        tonIdleWriteMetric(IN := FALSE, PT:= tIdleWriteMetric);
        GVL_MSG_XTS.MetricsMessageCtrl.Cmd                      := E_MESSAGE_CTRL.MSG_CTRL_NULL;
    END_CASE
END_CASE
//#################################################################################################################
//  Transport Metrics/
//#################################################################################################################
//#################################################################################################################
//#################################################################################################################

ACTION Init:
CASE eInit
OF
  E_PROGRESS.PROGRESS_INVALID:          // startup procedure for your application
    eInit                               := E_PROGRESS.PROGRESS_INIT;

  E_PROGRESS.PROGRESS_INIT:
      nProcess                                        := 1;
      tProcess[nProcess]                              := T#750MS;

      GVL_APPLICATION.Simulation[nProcess].HandshakeRoute:= E_PROCESS_HANDSHAKE.E_SHAKE_DOUBLE;

      GVL_APPLICATION.Simulation[nProcess].StationFirst  := 1;
      GVL_APPLICATION.Simulation[nProcess].StationLast   := 16;

      GVL_APPLICATION.Simulation[nProcess].TargetFirst   := 20;
      GVL_APPLICATION.Simulation[nProcess].TargetLast    := 35;
      GVL_APPLICATION.Simulation[nProcess].TargetMask    := 2#0001; // mask for target station

      GVL_APPLICATION.Simulation[nProcess].CheckRangeLow :=   10.0;
      GVL_APPLICATION.Simulation[nProcess].CheckRangeHigh:= 1600.0;

      //---------------------------------------------------------

      // 2

      //---------------------------------------------------------
      nProcess                                        := 3;
      tProcess[nProcess]                              := T#2400MS;

      GVL_APPLICATION.Simulation[nProcess].HandshakeRoute:= E_PROCESS_HANDSHAKE.E_SHAKE_DOUBLE;

      GVL_APPLICATION.Simulation[nProcess].StationFirst  := 20;
      GVL_APPLICATION.Simulation[nProcess].StationLast   := 35;

      GVL_APPLICATION.Simulation[nProcess].TargetFirst   := 37;
      GVL_APPLICATION.Simulation[nProcess].TargetLast    := 37;
      GVL_APPLICATION.Simulation[nProcess].TargetMask    := 2#0001; // mask for target station

      GVL_APPLICATION.Simulation[nProcess].CheckRangeLow := 9000.0;
      GVL_APPLICATION.Simulation[nProcess].CheckRangeHigh:= 12100.0;

      //---------------------------------------------------------
      nProcess                                        := 4;
      tProcess[nProcess]                              := T#0MS;

      GVL_APPLICATION.Simulation[nProcess].HandshakeRoute:= E_PROCESS_HANDSHAKE.E_SHAKE_SEND;

      GVL_APPLICATION.Simulation[nProcess].StationFirst  := 37;
      GVL_APPLICATION.Simulation[nProcess].StationLast   := 37;

      GVL_APPLICATION.Simulation[nProcess].TargetFirst   := 38;
      GVL_APPLICATION.Simulation[nProcess].TargetLast    := 38;
      GVL_APPLICATION.Simulation[nProcess].TargetMask    := 2#0001; // mask for target station

      GVL_APPLICATION.Simulation[nProcess].CheckRangeLow := 12850.0;
      GVL_APPLICATION.Simulation[nProcess].CheckRangeHigh:= 13000.0;

      //---------------------------------------------------------
      nProcess                                        := 5;
      tProcess[nProcess]                              := T#0MS;

      GVL_APPLICATION.Simulation[nProcess].HandshakeRoute:= E_PROCESS_HANDSHAKE.E_SHAKE_SEND;

      GVL_APPLICATION.Simulation[nProcess].StationFirst  := 38;
      GVL_APPLICATION.Simulation[nProcess].StationLast   := 38;

      GVL_APPLICATION.Simulation[nProcess].TargetFirst   := 39;
      GVL_APPLICATION.Simulation[nProcess].TargetLast    := 39;
      GVL_APPLICATION.Simulation[nProcess].TargetMask    := 2#0001; // mask for target station

      GVL_APPLICATION.Simulation[nProcess].CheckRangeLow := 13900.0;
      GVL_APPLICATION.Simulation[nProcess].CheckRangeHigh:= 14100.0;

      //---------------------------------------------------------
      nProcess                                        := 6;
      tProcess[nProcess]                              := T#0MS;

      GVL_APPLICATION.Simulation[nProcess].HandshakeRoute:= E_PROCESS_HANDSHAKE.E_SHAKE_SEND;

      GVL_APPLICATION.Simulation[nProcess].StationFirst  := 39;
      GVL_APPLICATION.Simulation[nProcess].StationLast   := 39;

      GVL_APPLICATION.Simulation[nProcess].TargetFirst   := 41;
      GVL_APPLICATION.Simulation[nProcess].TargetLast    := 52;
      GVL_APPLICATION.Simulation[nProcess].TargetMask    := 2#0001; // mask for target station

      GVL_APPLICATION.Simulation[nProcess].CheckRangeLow := 14200.0;
      GVL_APPLICATION.Simulation[nProcess].CheckRangeHigh:= 14400.0;

      //---------------------------------------------------------
      nProcess                                        := 7;
      tProcess[nProcess]                              := T#3200MS;

      GVL_APPLICATION.Simulation[nProcess].HandshakeRoute:= E_PROCESS_HANDSHAKE.E_SHAKE_FAST;

      GVL_APPLICATION.Simulation[nProcess].StationFirst  := 41;
      GVL_APPLICATION.Simulation[nProcess].StationLast   := 52;

      GVL_APPLICATION.Simulation[nProcess].TargetFirst   := 57;
      GVL_APPLICATION.Simulation[nProcess].TargetLast    := 57;
      GVL_APPLICATION.Simulation[nProcess].TargetMask    := 2#0001; // mask for target station

      GVL_APPLICATION.Simulation[nProcess].CheckRangeLow := 14400.0;
      GVL_APPLICATION.Simulation[nProcess].CheckRangeHigh:= 17000.0;

      //---------------------------------------------------------
      nProcess                                        := 8;
      tProcess[nProcess]                              := T#0MS;

      GVL_APPLICATION.Simulation[nProcess].HandshakeRoute:= E_PROCESS_HANDSHAKE.E_SHAKE_SEND;

      GVL_APPLICATION.Simulation[nProcess].StationFirst  := 57;
      GVL_APPLICATION.Simulation[nProcess].StationLast   := 57;

      GVL_APPLICATION.Simulation[nProcess].TargetFirst   := 58;
      GVL_APPLICATION.Simulation[nProcess].TargetLast    := 65;
      GVL_APPLICATION.Simulation[nProcess].TargetMask    := 2#0001; // mask for target station

      GVL_APPLICATION.Simulation[nProcess].CheckRangeLow := 17500.0;
      GVL_APPLICATION.Simulation[nProcess].CheckRangeHigh:= 18100.0;

      //---------------------------------------------------------
      nProcess                                        := 9;
      tProcess[nProcess]                              := T#3200MS;

      GVL_APPLICATION.Simulation[nProcess].HandshakeRoute:= E_PROCESS_HANDSHAKE.E_SHAKE_SINGLE;

      GVL_APPLICATION.Simulation[nProcess].StationFirst  := 58;
      GVL_APPLICATION.Simulation[nProcess].StationLast   := 65;

      GVL_APPLICATION.Simulation[nProcess].TargetFirst   := 70;
      GVL_APPLICATION.Simulation[nProcess].TargetLast    := 70;
      GVL_APPLICATION.Simulation[nProcess].TargetMask    := 2#0001; // mask for target station

      GVL_APPLICATION.Simulation[nProcess].CheckRangeLow := 19400.0;
      GVL_APPLICATION.Simulation[nProcess].CheckRangeHigh:= 20500.0;

      //---------------------------------------------------------
      nProcess                                        := 10;
      tProcess[nProcess]                              := T#0MS;

      GVL_APPLICATION.Simulation[nProcess].HandshakeRoute:= E_PROCESS_HANDSHAKE.E_SHAKE_SEND;

      GVL_APPLICATION.Simulation[nProcess].StationFirst  := 70;
      GVL_APPLICATION.Simulation[nProcess].StationLast   := 70;

      GVL_APPLICATION.Simulation[nProcess].TargetFirst   := 71;
      GVL_APPLICATION.Simulation[nProcess].TargetLast    := 82;
      GVL_APPLICATION.Simulation[nProcess].TargetMask    := 2#0001; // mask for target station

      GVL_APPLICATION.Simulation[nProcess].CheckRangeLow := 20600.0;
      GVL_APPLICATION.Simulation[nProcess].CheckRangeHigh:= 21400.0;

      //---------------------------------------------------------
      nProcess                                        := 12;
      tProcess[nProcess]                              := T#4600MS;

      GVL_APPLICATION.Simulation[nProcess].HandshakeRoute:= E_PROCESS_HANDSHAKE.E_SHAKE_DOUBLE;

      GVL_APPLICATION.Simulation[nProcess].StationFirst  := 71;
      GVL_APPLICATION.Simulation[nProcess].StationLast   := 82;

      GVL_APPLICATION.Simulation[nProcess].TargetFirst   := 91;
      GVL_APPLICATION.Simulation[nProcess].TargetLast    := 91;
      GVL_APPLICATION.Simulation[nProcess].TargetMask    := 2#0001; // mask for target station

      GVL_APPLICATION.Simulation[nProcess].CheckRangeLow := 21400.0;
      GVL_APPLICATION.Simulation[nProcess].CheckRangeHigh:= 22800.0;

      //---------------------------------------------------------
      nProcess                                        := 13;
      tProcess[nProcess]                              := T#00MS;

      GVL_APPLICATION.Simulation[nProcess].HandshakeRoute:= E_PROCESS_HANDSHAKE.E_SHAKE_SEND;

      GVL_APPLICATION.Simulation[nProcess].StationFirst  := 91;
      GVL_APPLICATION.Simulation[nProcess].StationLast   := 91;

      GVL_APPLICATION.Simulation[nProcess].TargetFirst   := 95;
      GVL_APPLICATION.Simulation[nProcess].TargetLast    := 95;
      GVL_APPLICATION.Simulation[nProcess].TargetMask    := 2#0001; // mask for target station

      GVL_APPLICATION.Simulation[nProcess].CheckRangeLow := 22800.0;
      GVL_APPLICATION.Simulation[nProcess].CheckRangeHigh:= 23500.0;

      //---------------------------------------------------------
      nProcess                                        := 14;
      tProcess[nProcess]                              := T#0MS;

      GVL_APPLICATION.Simulation[nProcess].HandshakeRoute:= E_PROCESS_HANDSHAKE.E_SHAKE_SEND;

      GVL_APPLICATION.Simulation[nProcess].StationFirst  := 95;
      GVL_APPLICATION.Simulation[nProcess].StationLast   := 95;

      GVL_APPLICATION.Simulation[nProcess].TargetFirst   := 120;
      GVL_APPLICATION.Simulation[nProcess].TargetLast    := 133;
      GVL_APPLICATION.Simulation[nProcess].TargetMask    := 2#0001; // mask for target station

      GVL_APPLICATION.Simulation[nProcess].CheckRangeLow := 24000.0;
      GVL_APPLICATION.Simulation[nProcess].CheckRangeHigh:= 24100.0;

      //---------------------------------------------------------
      nProcess                                        := 15;
      tProcess[nProcess]                              := T#2500MS;

      GVL_APPLICATION.Simulation[nProcess].HandshakeRoute:= E_PROCESS_HANDSHAKE.E_SHAKE_DOUBLE;

      GVL_APPLICATION.Simulation[nProcess].StationFirst  := 120;
      GVL_APPLICATION.Simulation[nProcess].StationLast   := 133;

      GVL_APPLICATION.Simulation[nProcess].TargetFirst   := 140;
      GVL_APPLICATION.Simulation[nProcess].TargetLast    := 140;
      GVL_APPLICATION.Simulation[nProcess].TargetMask    := 2#0001; // mask for target station

      GVL_APPLICATION.Simulation[nProcess].CheckRangeLow := 24200.0;
      GVL_APPLICATION.Simulation[nProcess].CheckRangeHigh:= 27500.0;

      //---------------------------------------------------------
      nProcess                                        := 16;
      tProcess[nProcess]                              := T#0MS;

      GVL_APPLICATION.Simulation[nProcess].HandshakeRoute:= E_PROCESS_HANDSHAKE.E_SHAKE_SEND;

      GVL_APPLICATION.Simulation[nProcess].StationFirst  := 140;
      GVL_APPLICATION.Simulation[nProcess].StationLast   := 140;

      GVL_APPLICATION.Simulation[nProcess].TargetFirst   := 141;
      GVL_APPLICATION.Simulation[nProcess].TargetLast    := 141;
      GVL_APPLICATION.Simulation[nProcess].TargetMask    := 2#0001; // mask for target station

      GVL_APPLICATION.Simulation[nProcess].CheckRangeLow := 27970.0;
      GVL_APPLICATION.Simulation[nProcess].CheckRangeHigh:= 1250.0;

      //---------------------------------------------------------
      nProcess                                        := 17;
      tProcess[nProcess]                              := T#0MS;

      GVL_APPLICATION.Simulation[nProcess].HandshakeRoute:= E_PROCESS_HANDSHAKE.E_SHAKE_SEND;

      GVL_APPLICATION.Simulation[nProcess].StationFirst  := 141;
      GVL_APPLICATION.Simulation[nProcess].StationLast   := 141;

      GVL_APPLICATION.Simulation[nProcess].TargetFirst   := 142;
      GVL_APPLICATION.Simulation[nProcess].TargetLast    := 142;
      GVL_APPLICATION.Simulation[nProcess].TargetMask    := 2#0001; // mask for target station

      GVL_APPLICATION.Simulation[nProcess].CheckRangeLow := 3950.0;
      GVL_APPLICATION.Simulation[nProcess].CheckRangeHigh:= 4100.0;

      //---------------------------------------------------------
      nProcess                                        := 18;
      tProcess[nProcess]                              := T#0MS;

      GVL_APPLICATION.Simulation[nProcess].HandshakeRoute:= E_PROCESS_HANDSHAKE.E_SHAKE_SEND;

      GVL_APPLICATION.Simulation[nProcess].StationFirst  := 142;
      GVL_APPLICATION.Simulation[nProcess].StationLast   := 142;

      GVL_APPLICATION.Simulation[nProcess].TargetFirst   := 20;
      GVL_APPLICATION.Simulation[nProcess].TargetLast    := 35;
      GVL_APPLICATION.Simulation[nProcess].TargetMask    := 2#0001; // mask for target station

      GVL_APPLICATION.Simulation[nProcess].CheckRangeLow := 4500.0;
      GVL_APPLICATION.Simulation[nProcess].CheckRangeHigh:= 5600.0;


    eInit                                                 := E_PROGRESS.PROGRESS_BUSY;

  E_PROGRESS.PROGRESS_BUSY:
    GVL_MSG_XTS.TransportMessageCtrl.Cmd                  := E_MESSAGE_CTRL.MSG_CTRL_INIT;
    GVL_MSG_XTS.MetricsMessageCtrl.Cmd                    := E_MESSAGE_CTRL.MSG_CTRL_INIT;
    eInit                                                 := E_PROGRESS.PROGRESS_PREPARE;

  E_PROGRESS.PROGRESS_PREPARE:
    eInit                                                 := E_PROGRESS.PROGRESS_STARTUP;

  E_PROGRESS.PROGRESS_STARTUP:
    eInit                                                 := E_PROGRESS.PROGRESS_DONE;
    FOR nProcess := 1 TO MAX_PROCESS
    DO
      IF (GVL_APPLICATION.Simulation[nProcess].StationCount > 0)
      THEN
        GVL_APPLICATION.Simulation[nProcess].EnableProcess := TO_DWORD(EXPT(2,GVL_APPLICATION.Simulation[nProcess].StationCount))-1;
        GVL_APPLICATION.Simulation[nProcess].MoverEnter    := TRUE;
        GVL_APPLICATION.Simulation[nProcess].MoverOut      := TRUE;

      END_IF
    END_FOR
END_CASE
END_ACTION

END_PROGRAM

(* stored: Version 1.1.0.1
   POU MAIN_APP: Id {aed82ec5-7c0f-4ed8-9d95-00008ab7747f}, SpecialFunc None
   Action Init: Id {69838e0d-19cf-48fe-8b42-ee1af1eba2b6} *)
